{attribute 'linkalways'}
{attribute 'no_explicit_call' := 'Use the methods of this class'}
{attribute 'enable_dynamic_creation'}
FUNCTION_BLOCK Gyro_Simulated IMPLEMENTS I_Gyro
VAR
	link : REFERENCE TO SimulatorLink;
END_VAR

METHOD FB_init : BOOL
VAR_INPUT
	bInitRetains : BOOL;
	bInCopyCode : BOOL;
	simulator : REFERENCE TO SimulatorLink;
END_VAR
link REF= simulator;
END_METHOD

METHOD StartBiasCalibration
// The simulated gyro has no calibration of its own. Bias is estimated in HeadingFusion.
END_METHOD

PROPERTY YawRateInRadPerS : LREAL
GET
YawRateInRadPerS := SimulatorIo.feedback.angularRateInRadPerS.z;
END_GET
END_PROPERTY

PROPERTY AngularRateInRadPerS : Vector3
GET
AngularRateInRadPerS := SimulatorIo.feedback.angularRateInRadPerS;
END_GET
END_PROPERTY

PROPERTY TimestampInNs : ULINT
GET
TimestampInNs := SimulatorIo.feedback.timeInNs;
END_GET
END_PROPERTY

PROPERTY IsValid : BOOL
GET
IsValid := __ISVALIDREF(link) AND_THEN link.IsConnected;
END_GET
END_PROPERTY

END_FUNCTION_BLOCK

(* stored: Version 1.1.0.1, ProductVersion 3.1.4026.12
   POU Gyro_Simulated: Id {4514b4b8-d81e-559f-97c2-245e28b90dbd}, SpecialFunc None
   Method FB_init: Id {576750ad-b360-5306-b633-18829c7c943a}
   Method StartBiasCalibration: Id {a9e518d6-8ef0-5b9a-b66a-c86cdd4b5b62}
   Property YawRateInRadPerS: Id {6b8f2a0b-ed68-5a9b-95c6-c7e6ab0ab276}
   Get Get: Id {bef85936-34ad-5498-81c2-ef0e5b7a88a0}
   Property AngularRateInRadPerS: Id {5c71fdd9-2b7c-5963-bca3-c500b1b3304c}
   Get Get: Id {7861b59a-a0a0-5460-96e1-08b09760ed98}
   Property TimestampInNs: Id {719c20c0-1047-5d5f-ac84-ede0bf00fd8a}
   Get Get: Id {8cc0bfd1-f9c2-5741-907c-d08b5ca383b0}
   Property IsValid: Id {5e8d67d2-6198-57c5-ba2d-3450b85e5bec}
   Get Get: Id {8d2806f6-a03d-5243-849f-b5ae1f51b6e5} *)
